(* IEC 61131-3 sources: llm-plc-st-eval/data/processed_definitivo/gemini-3.1-pro-preview/A1/few_shot, 3 files *)

(* ---- ejec_1.st ---- *)
FUNCTION_BLOCK FB_PID
VAR_INPUT
    SP : REAL; (* Consigna *)
    PV : REAL; (* Variable de proceso *)
    Kp : REAL; (* Ganancia proporcional *)
    Ti : REAL; (* Tiempo integral en segundos *)
    Td : REAL; (* Tiempo derivativo en segundos *)
    ciclo : TIME; (* Periodo de muestreo *)
END_VAR
VAR_OUTPUT
    CV : REAL; (* Variable de control (0.0 a 100.0) *)
END_VAR
VAR
    e : REAL; (* Error actual *)
    e_prev : REAL; (* Error del ciclo anterior *)
    integral_acc : REAL; (* Acumulador de la integral del error *)
    dt_sec : REAL; (* Tiempo de ciclo en segundos *)
    deriv : REAL; (* Derivada del error *)
    I_term : REAL; (* Termino integral *)
    D_term : REAL; (* Termino derivativo *)
    CV_temp : REAL; (* Variable de control sin limitar *)
END_VAR

(* Conversion del tiempo de ciclo a segundos *)
dt_sec := TIME_TO_REAL(ciclo) / 1000.0;

(* Calculo del error *)
e := SP - PV;

(* Accion Integral con Anti-windup por clamping *)
IF Ti > 0.0 THEN
    (* Evita acumular error positivo si CV esta al 100%, o negativo si CV esta al 0% *)
    IF NOT ((CV >= 100.0 AND e > 0.0) OR (CV <= 0.0 AND e < 0.0)) THEN
        integral_acc := integral_acc + (e * dt_sec);
    END_IF;
    I_term := integral_acc / Ti;
ELSE
    integral_acc := 0.0;
    I_term := 0.0;
END_IF;

(* Accion Derivativa *)
IF dt_sec > 0.0 THEN
    deriv := (e - e_prev) / dt_sec;
ELSE
    deriv := 0.0;
END_IF;
D_term := Td * deriv;

(* Ecuacion PID estandar *)
CV_temp := Kp * (e + I_term + D_term);

(* Limitacion de la salida (0.0 a 100.0) *)
IF CV_temp > 100.0 THEN
    CV := 100.0;
ELSIF CV_temp < 0.0 THEN
    CV := 0.0;
ELSE
    CV := CV_temp;
END_IF;

(* Actualizacion del error para el calculo derivativo del proximo ciclo *)
e_prev := e;

END_FUNCTION_BLOCK

(* ---- ejec_2.st ---- *)
FUNCTION_BLOCK FB_PID
VAR_INPUT
    SP : REAL; (* Consigna *)
    PV : REAL; (* Variable de proceso *)
    Kp : REAL; (* Ganancia proporcional *)
    Ti : REAL; (* Tiempo integral en segundos *)
    Td : REAL; (* Tiempo derivativo en segundos *)
    ciclo : TIME; (* Periodo de muestreo *)
END_VAR
VAR_OUTPUT
    CV : REAL; (* Porcentaje de mando (0.0 a 100.0) *)
END_VAR
VAR
    e : REAL; (* Error actual *)
    e_prev : REAL; (* Error del ciclo anterior *)
    integral : REAL; (* Acumulador de la integral *)
    derivada : REAL; (* Tasa de cambio del error *)
    dt : REAL; (* Tiempo de ciclo en segundos *)
    CV_raw : REAL; (* Salida calculada sin limitar *)
END_VAR

(* Conversion del tiempo de ciclo a segundos *)
dt := DINT_TO_REAL(TIME_TO_DINT(ciclo)) / 1000.0;

IF dt > 0.0 THEN
    (* Calculo del error *)
    e := SP - PV;

    (* Accion integral con anti-windup por clamping *)
    IF Ti > 0.0 THEN
        (* Evitar integracion si la salida esta saturada y el error empuja en la misma direccion *)
        IF NOT ((CV >= 100.0 AND e > 0.0) OR (CV <= 0.0 AND e < 0.0)) THEN
            integral := integral + (e * dt);
        END_IF;
    ELSE
        integral := 0.0; (* Desactivar accion integral si Ti <= 0.0 *)
    END_IF;

    (* Accion derivativa sobre el error *)
    derivada := (e - e_prev) / dt;

    (* Calculo de la salida (Forma estandar del PID) *)
    IF Ti > 0.0 THEN
        CV_raw := Kp * (e + (integral / Ti) + (Td * derivada));
    ELSE
        CV_raw := Kp * (e + (Td * derivada));
    END_IF;

    (* Limitacion de la salida al rango 0.0 - 100.0 *)
    IF CV_raw > 100.0 THEN
        CV := 100.0;
    ELSIF CV_raw < 0.0 THEN
        CV := 0.0;
    ELSE
        CV := CV_raw;
    END_IF;

    (* Actualizar el error anterior para el proximo ciclo *)
    e_prev := e;
END_IF;
END_FUNCTION_BLOCK

(* ---- ejec_3.st ---- *)
FUNCTION_BLOCK FB_PID
VAR_INPUT
    SP : REAL; (* Consigna *)
    PV : REAL; (* Variable de proceso *)
    Kp : REAL; (* Ganancia proporcional *)
    Ti : REAL; (* Tiempo integral en segundos *)
    Td : REAL; (* Tiempo derivativo en segundos *)
    ciclo : TIME; (* Periodo de muestreo *)
END_VAR
VAR_OUTPUT
    CV : REAL; (* Porcentaje de mando (0.0 a 100.0) *)
END_VAR
VAR
    e : REAL; (* Error actual *)
    e_prev : REAL; (* Error del ciclo anterior *)
    integral : REAL; (* Acumulador de la integral del error *)
    dt : REAL; (* Tiempo de ciclo en segundos *)
    P_term : REAL; (* Accion proporcional *)
    I_term : REAL; (* Accion integral *)
    D_term : REAL; (* Accion derivativa *)
    CV_unc : REAL; (* Salida calculada sin limitar *)
END_VAR

(* Conversion del tiempo de ciclo a segundos *)
dt := TIME_TO_REAL(ciclo) / 1000.0;
IF dt <= 0.0 THEN
    dt := 0.001; (* Evitar division por cero *)
END_IF;

(* Calculo del error *)
e := SP - PV;

(* Accion proporcional *)
P_term := Kp * e;

(* Accion derivativa sobre el error *)
D_term := Kp * Td * ((e - e_prev) / dt);

(* Accion integral y calculo de salida sin limitar *)
IF Ti > 0.0 THEN
    (* Se evalua con la integral tentativa para el ciclo actual *)
    I_term := Kp * ((integral + (e * dt)) / Ti);
ELSE
    I_term := 0.0;
    integral := 0.0;
END_IF;

CV_unc := P_term + I_term + D_term;

(* Anti-windup por clamping: actualizacion del acumulador integral *)
IF Ti > 0.0 THEN
    (* No acumula si esta saturado al maximo y el error es positivo, o saturado al minimo y el error es negativo *)
    IF NOT ((CV_unc >= 100.0 AND e > 0.0) OR (CV_unc <= 0.0 AND e < 0.0)) THEN
        integral := integral + (e * dt);
    END_IF;
END_IF;

(* Limitacion de la salida CV al rango 0.0 - 100.0 *)
IF CV_unc > 100.0 THEN
    CV := 100.0;
ELSIF CV_unc < 0.0 THEN
    CV := 0.0;
ELSE
    CV := CV_unc;
END_IF;

(* Memoria del error para la derivada en el proximo ciclo *)
e_prev := e;
END_FUNCTION_BLOCK
